Fanuc KAREL source: KA00096.KL

PROGRAM KA00096
%NOLOCKGROUP
VAR
  SRC: JOINTPOS
  DST: ARRAY[2] OF SHORT
BEGIN
  DST[1] = SRC
END KA00096
